// TIA Portal V21 export
// export: Created 2026-10-12T12:46:19.0179761Z, ExportSetting WithDefaults, DisplayName Totally Integrated Automation Portal, DisplayVersion V21, DisplayName STEP 7 Professional, DisplayVersion V21, DisplayName STEP 7 Safety, DisplayVersion V21, DisplayName Tech WebApplication, DisplayVersion V21, DisplayName WinCC Basic/Comfort/Advanced, DisplayVersion V21, DisplayName WinCC Unified, DisplayVersion V21
TextList "AUTO STATUS"  ListRange=Decimal
  TextListEntry   EntryType=SingleValue, From=10, To=10, Text="AUTO RUNNING"
  TextListEntry   EntryType=SingleValue, From=20, To=20, Text="STOPPED"
  TextListEntry   EntryType=SingleValue, From=30, To=30, Text="WAITING FOR CAMERA ACK"
